// TIA Portal V21 export
// export: Created 2026-05-12T00:00:00.0000000Z, ExportSetting None
DATA_BLOCK "DB_HMI_Interface"   // DB200
{ S7_Optimized_Access := 'FALSE' }
   VAR
      Enabled : Bool := false;
      DefaultInt : Int;
      "电机/运行%2F" : Bool := true;
      Motor : Struct
         Config : Struct
            Speed : Real := 1.5;
         END_STRUCT;
      END_STRUCT;
      Samples : Array[0..1] of Int;
      Locked : Int := 7;
      Inherited : Struct
         Value : Int;
      END_STRUCT;
      LockedValue : Int := 9;
      Typed : "MotorType";
      Clock : DTL;
   END_VAR
BEGIN
   Samples[0] := 3;
END_DATA_BLOCK
